// TIA Portal V21 export
FUNCTION_BLOCK "Timed"   // FB30, GRAPH
TITLE = Timed carriage
// A carriage that runs and brakes, with step times: the defaults, both set, and only the maximum set.
   VAR_INPUT
      ACK_EF : Bool;
      go : Bool;
      arrived : Bool;
      stopped : Bool;
      jammed : Bool;
   END_VAR
   VAR_OUTPUT
      motor : Bool;
      brake : Bool;
   END_VAR
BEGIN
// Sequence
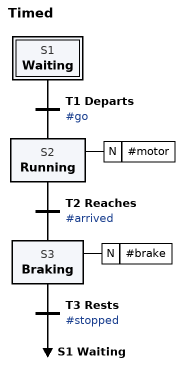
   // sequencer 1
   INITIAL_STEP Waiting:   // S1
   END_STEP
   TRANSITION Departs FROM Waiting TO Running   // T1
      := #go;
   END_TRANSITION
   STEP Running:   // S2, max time T#30S, warning time T#20S
      supervision V := #jammed;
              N    #motor
   END_STEP
   TRANSITION Reaches FROM Running TO Braking   // T2
      := #arrived;
   END_TRANSITION
   STEP Braking:   // S3, max time T#1M30S
              N    #brake
   END_STEP
   TRANSITION Rests FROM Braking TO Waiting   // T3, jump
      := #stopped;
   END_TRANSITION
END_FUNCTION_BLOCK
